DATA_BLOCK "FRK_HealthDefaults"
{ S7_Optimized_Access := 'TRUE' }
VERSION : 0.1
NON_RETAIN
VAR
    Config {ExternalAccessible := 'False'; ExternalVisible := 'False'; ExternalWritable := 'False'} : "ST_SystemHealthParCfg";
END_VAR
BEGIN
END_DATA_BLOCK
